SUBAPPLICATION logiBUS_AI_Calibrate_2P_OPC (* logiBUS_AI 2-Punkt-Kalibrierung, INI-persistiert, CO/CS per Methode, alles per OPC-UA (ohne VT) *)
  (* Standard: 61499-2; Description: Copyright (c) 2026 Meisterschulen am Ostbahnhof This program and the accompanying materials are made available under the terms of the Eclipse Public License 2.0 which is available at https://www.eclipse.org/legal/epl-2.0/ SPDX-License-Identifier: EPL-2.0 *)
  (* Version 1.1, 2026-11-25, Franz Höpfinger, Meisterschulen am Ostbahnhof, SERVER_0 -> MyLib::net::SERVER_0_QO (IND nur bei QO=TRUE, RSP intern). Ein gescheitertes RSP meldet IND mit QO=FALSE, direkt IND->RSP ergab eine Endlosschleife. *)
  (* Version 1.0, 2026-10-28, Franz Höpfinger, Meisterschulen am Ostbahnhof, Kopie von MyLib::sys::logiBUS_AI_Calibrate_2P_IDA_OPC v1.12 ohne VT, fuer Stationen ohne VT (keine isobus_UT-Libs). InputRaw -> MyLib::sys::logiBUS_AI_Raw_AR_OPC, Y_OFFSET_LIT/Y_SCALE_LIT -> MyLib::sys::OPC_TO_AR2, TriggerCO/CS -> SERVER_0 (IND->RSP), Publish* -> MyLib::sys::AR_TO_Publish_OPC. VT-Objekt-Parameter entfallen, Kalibrierlogik und INI-Keys unveraendert. *)
  PACKAGE MyLib::sys;
  IMPORT logiBUS::io::AI::logiBUS_AI;
  IMPORT logiBUS::io::AI::logiBUS_AI_S;
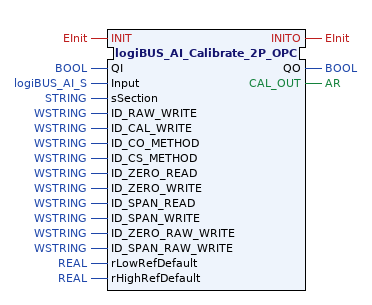
  EVENT_INPUT
    INIT : EInit; (* Initialization Request *)
  END_EVENT
  EVENT_OUTPUT
    INITO : EInit; (* Initialization Confirm *)
  END_EVENT
  VAR_INPUT
    QI : BOOL := TRUE; (* Quality Input - TRUE to enable service *)
    Input : logiBUS::io::AI::logiBUS_AI_S := logiBUS_AI::Invalid; (* Identify the Input AnalogInput_I1..I8 *)
    sSection : STRING; (* INI-Sektionsname fuer OFFSET/SCALE-Persistenz - pro Kanal eindeutig (z.B. 'AI_Calibrate_I1'), sonst kollidieren die Kanaele in settings.ini *)
    ID_RAW_WRITE : WSTRING; (* Rohwert-Ruckmelde-Adresse (DWORD 0-4095, ACTION=PUBLISH) *)
    ID_CAL_WRITE : WSTRING; (* Kalibrierter-Wert-Ruckmelde-Adresse (REAL, ACTION=PUBLISH) *)
    ID_CO_METHOD : WSTRING; (* Methodenadresse (CREATE_METHOD) fuer den CO-Trigger (Dashboard oder CLIENT_0 von STG1) *)
    ID_CS_METHOD : WSTRING; (* Methodenadresse (ACTION=CREATE_METHOD) fuer den argumentlosen CS-Trigger - siehe ID_CO_METHOD *)
    ID_ZERO_READ : WSTRING; (* Remote-Subscribe-Adresse ZERO-Referenzwert (REAL, ACTION=SUBSCRIBE) *)
    ID_ZERO_WRITE : WSTRING; (* Remote-Echo-Adresse ZERO-Referenzwert (REAL, ACTION=PUBLISH) *)
    ID_SPAN_READ : WSTRING; (* Remote-Subscribe-Adresse SPAN-Referenzwert (REAL, ACTION=SUBSCRIBE) *)
    ID_SPAN_WRITE : WSTRING; (* Remote-Echo-Adresse SPAN-Referenzwert (REAL, ACTION=PUBLISH) *)
    ID_ZERO_RAW_WRITE : WSTRING; (* Rohwert-am-ZERO-Kalibrierpunkt-Publish-Adresse (REAL, ACTION=PUBLISH) *)
    ID_SPAN_RAW_WRITE : WSTRING; (* Rohwert-am-SPAN-Kalibrierpunkt-Publish-Adresse (REAL, ACTION=PUBLISH) *)
    rLowRefDefault : REAL := REAL#0.0; (* Erstinbetriebnahme-Standardwert LOW_REF (INI_LOW_REF.DEFAULT_VALUE), bevor der Bediener selbst kalibriert - Fuellband/die meisten Sensoren: 0.0 *)
    rHighRefDefault : REAL := REAL#100.0; (* Erstinbetriebnahme-Standardwert HIGH_REF (INI_HIGH_REF.DEFAULT_VALUE), bevor der Bediener selbst kalibriert - z.B. 250.0 fuer Druck (0-250bar), 100.0 fuer Fuellband-Winkel (Prozent) *)
  END_VAR
  VAR_OUTPUT
    QO : BOOL; (* Quality Output - TRUE if service executed successfully *)
  END_VAR
  PLUGS
    CAL_OUT : adapter::types::unidirectional::AR; (* Kalibrierter Wert, lokal (= CALIBRATE.Y) - fuer Weiterverarbeitung auf derselben Station ohne OPC-UA-Roundtrip *)
  END_PLUGS
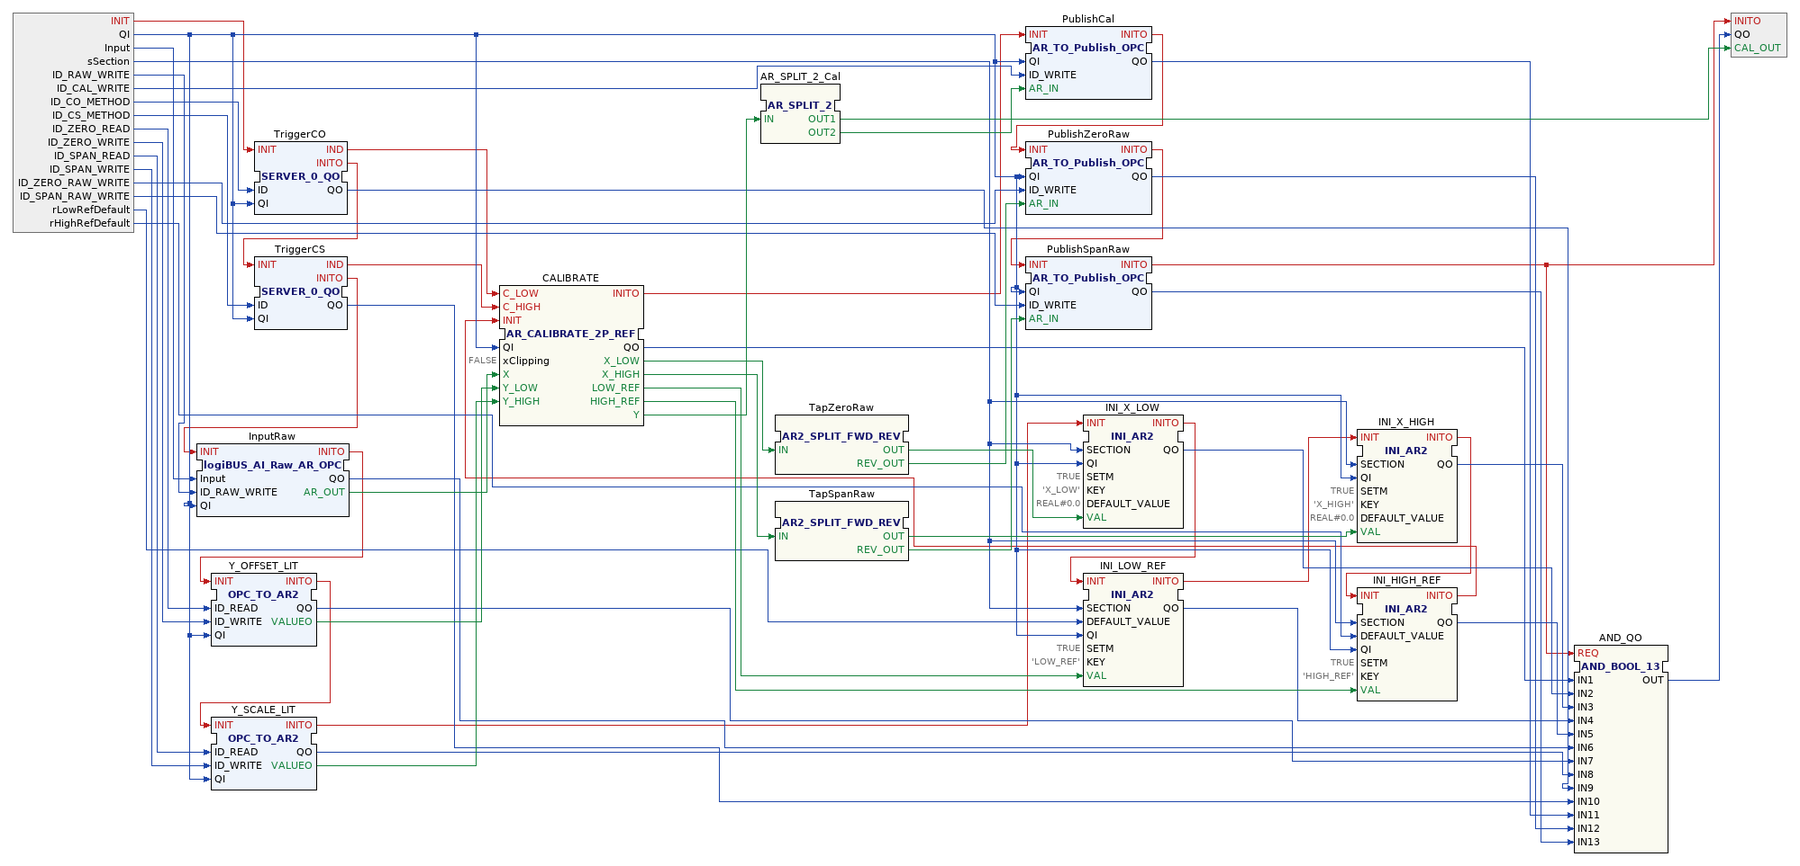
  (* INIT-Reihenfolge: INI-Werte (X_LOW/LOW_REF/X_HIGH/HIGH_REF) VOR CALIBRATE, sonst rechnet CALIBRATE beim Start kurz mit 0-Kalibrierpunkten. *)
  FBS
    CALIBRATE : adapter::Engineering::measurements::AR_CALIBRATE_2P_REF(xClipping := FALSE);
    INI_X_LOW : eclipse4diac::storage::INI_AR2(SETM := TRUE, KEY := 'X_LOW', DEFAULT_VALUE := REAL#0.0);
    INI_X_HIGH : eclipse4diac::storage::INI_AR2(SETM := TRUE, KEY := 'X_HIGH', DEFAULT_VALUE := REAL#0.0);
    INI_LOW_REF : eclipse4diac::storage::INI_AR2(SETM := TRUE, KEY := 'LOW_REF');
    INI_HIGH_REF : eclipse4diac::storage::INI_AR2(SETM := TRUE, KEY := 'HIGH_REF');
    TapZeroRaw : adapter::events::bidirectional::AR2_SPLIT_FWD_REV;
    TapSpanRaw : adapter::events::bidirectional::AR2_SPLIT_FWD_REV;
    AR_SPLIT_2_Cal : adapter::events::unidirectional::AR_SPLIT_2;
    AND_QO : iec61131::booleanOperators::AND_BOOL_13;
  END_FBS
  SUBAPPS
    InputRaw : MyLib::sys::logiBUS_AI_Raw_AR_OPC;
    Y_OFFSET_LIT : MyLib::sys::OPC_TO_AR2;
    Y_SCALE_LIT : MyLib::sys::OPC_TO_AR2;
    TriggerCO : MyLib::net::SERVER_0_QO; (* RSP direkt auf IND (sonst 4s Server-Lock) *)
    TriggerCS : MyLib::net::SERVER_0_QO; (* RSP direkt auf IND (sonst 4s Server-Lock) *)
    PublishCal : MyLib::sys::AR_TO_Publish_OPC;
    PublishZeroRaw : MyLib::sys::AR_TO_Publish_OPC;
    PublishSpanRaw : MyLib::sys::AR_TO_Publish_OPC;
  END_SUBAPPS
  EVENT_CONNECTIONS
    TriggerCO.IND TO CALIBRATE.C_LOW;
    TriggerCS.IND TO CALIBRATE.C_HIGH;
    CALIBRATE.INITO TO PublishCal.INIT;
    InputRaw.INITO TO Y_OFFSET_LIT.INIT;
    Y_OFFSET_LIT.INITO TO Y_SCALE_LIT.INIT;
    TriggerCO.INITO TO TriggerCS.INIT;
    PublishCal.INITO TO PublishZeroRaw.INIT;
    PublishZeroRaw.INITO TO PublishSpanRaw.INIT;
    INIT TO TriggerCO.INIT;
    TriggerCS.INITO TO InputRaw.INIT;
    Y_SCALE_LIT.INITO TO INI_X_LOW.INIT;
    INI_HIGH_REF.INITO TO CALIBRATE.INIT;
    INI_X_LOW.INITO TO INI_LOW_REF.INIT;
    INI_LOW_REF.INITO TO INI_X_HIGH.INIT;
    INI_X_HIGH.INITO TO INI_HIGH_REF.INIT;
    PublishSpanRaw.INITO TO AND_QO.REQ;
    PublishSpanRaw.INITO TO INITO;
  END_CONNECTIONS
  DATA_CONNECTIONS
    Input TO InputRaw.Input;
    sSection TO INI_X_LOW.SECTION;
    sSection TO INI_X_HIGH.SECTION;
    sSection TO INI_LOW_REF.SECTION;
    sSection TO INI_HIGH_REF.SECTION;
    rLowRefDefault TO INI_LOW_REF.DEFAULT_VALUE;
    rHighRefDefault TO INI_HIGH_REF.DEFAULT_VALUE;
    ID_RAW_WRITE TO InputRaw.ID_RAW_WRITE;
    ID_CAL_WRITE TO PublishCal.ID_WRITE;
    ID_CO_METHOD TO TriggerCO.ID;
    ID_CS_METHOD TO TriggerCS.ID;
    ID_ZERO_READ TO Y_OFFSET_LIT.ID_READ;
    ID_ZERO_WRITE TO Y_OFFSET_LIT.ID_WRITE;
    ID_SPAN_READ TO Y_SCALE_LIT.ID_READ;
    ID_SPAN_WRITE TO Y_SCALE_LIT.ID_WRITE;
    ID_ZERO_RAW_WRITE TO PublishZeroRaw.ID_WRITE;
    ID_SPAN_RAW_WRITE TO PublishSpanRaw.ID_WRITE;
    QI TO CALIBRATE.QI;
    QI TO INI_X_LOW.QI;
    QI TO INI_X_HIGH.QI;
    QI TO INI_LOW_REF.QI;
    QI TO INI_HIGH_REF.QI;
    QI TO InputRaw.QI;
    QI TO Y_OFFSET_LIT.QI;
    QI TO Y_SCALE_LIT.QI;
    QI TO TriggerCO.QI;
    QI TO TriggerCS.QI;
    QI TO PublishCal.QI;
    QI TO PublishZeroRaw.QI;
    QI TO PublishSpanRaw.QI;
    CALIBRATE.QO TO AND_QO.IN1;
    INI_X_LOW.QO TO AND_QO.IN2;
    INI_X_HIGH.QO TO AND_QO.IN3;
    INI_LOW_REF.QO TO AND_QO.IN4;
    INI_HIGH_REF.QO TO AND_QO.IN5;
    InputRaw.QO TO AND_QO.IN6;
    Y_OFFSET_LIT.QO TO AND_QO.IN7;
    Y_SCALE_LIT.QO TO AND_QO.IN8;
    TriggerCO.QO TO AND_QO.IN9;
    TriggerCS.QO TO AND_QO.IN10;
    PublishCal.QO TO AND_QO.IN11;
    PublishZeroRaw.QO TO AND_QO.IN12;
    PublishSpanRaw.QO TO AND_QO.IN13;
    AND_QO.OUT TO QO;
  END_CONNECTIONS
  ADAPTER_CONNECTIONS
    InputRaw.AR_OUT TO CALIBRATE.X;
    CALIBRATE.X_LOW TO TapZeroRaw.IN;
    TapZeroRaw.OUT TO INI_X_LOW.VAL;
    TapZeroRaw.REV_OUT TO PublishZeroRaw.AR_IN;
    CALIBRATE.X_HIGH TO TapSpanRaw.IN;
    TapSpanRaw.OUT TO INI_X_HIGH.VAL;
    TapSpanRaw.REV_OUT TO PublishSpanRaw.AR_IN;
    CALIBRATE.LOW_REF TO INI_LOW_REF.VAL;
    CALIBRATE.HIGH_REF TO INI_HIGH_REF.VAL;
    Y_OFFSET_LIT.VALUEO TO CALIBRATE.Y_LOW;
    Y_SCALE_LIT.VALUEO TO CALIBRATE.Y_HIGH;
    CALIBRATE.Y TO AR_SPLIT_2_Cal.IN;
    AR_SPLIT_2_Cal.OUT1 TO CAL_OUT;
    AR_SPLIT_2_Cal.OUT2 TO PublishCal.AR_IN;
  END_CONNECTIONS
END_SUBAPPLICATION
